TYPE ST_PolarIIChamber_ServiceCtrl :
STRUCT
	Chamber : ST_PolarIIChamber_ChamberServiceCtrl;
	Arm : ARRAY[1..4] OF ST_PolarIIChamber_ArmServiceCtrl;
	Cup : ARRAY[1..4] OF ST_PolarIIChamber_CupServiceCtrl;
	Holder : ST_PolarIIChamber_HolderServiceCtrl;
	FixedNozzle : ARRAY[1..4] OF ST_PolarIIChamber_NozzleSupplyServiceCtrl;
	OutsideRing : ST_PolarIIChamber_OutsideRingServiceCtrl;
	Shutter : ST_PolarIIChamber_OpenCloseServiceCtrl;
	Exhaust : ST_PolarIIChamber_ExhaustServiceCtrl;
	SideVent : ARRAY[1..4] OF ST_PolarIIChamber_OpenCloseServiceCtrl;
END_STRUCT
END_TYPE

(* stored: Version 1.1.0.1, ProductVersion 3.1.4026.18
   DUT ST_PolarIIChamber_ServiceCtrl: Id {14000000-0000-0000-0000-000000000073} *)
